Fanuc KAREL source: KT00666.KL

PROGRAM KT00666
%NOLOCKGROUP
VAR
  P1: XYZWPR
  P2: XYZWPR
  OUT: BOOLEAN
BEGIN
  P1.X = 1.0
  P2.Y = 2.0
  P1.X = 1.0
  P2.Y = 2.0
  OUT = + P1
END KT00666
